// Objet Sécurités : la station (ou la machine) lit l'état de ses circuits (docs/03 § 8.2, docs/05 § 4.2)
INTERFACE I_SafetyCircuits

PROPERTY AllOk : BOOL
GET
END_GET
END_PROPERTY

END_INTERFACE

(* stored: Version 1.1.0.1, ProductVersion 3.1.4024.12
   Itf I_SafetyCircuits: Id {5163598b-a23b-597a-8474-79c1a183c996}
   Property AllOk: Id {f8bd1ace-d4d0-57b5-ad8b-001d4f8ae3cc}
   Get Get: Id {27a4d94e-7cd6-520f-a379-53e88db2f075} *)
